FUNCTION SPEED_CONTROL : INT
VAR_INPUT
	ixLevel : INT;
END_VAR

SPEED_CONTROL := (50 - ixLevel) * 10;
IF SPEED_CONTROL < 0 THEN;
	SPEED_CONTROL := 0;
END_IF

END_FUNCTION

(* stored: Version 1.1.0.1
   POU SPEED_CONTROL: Id {2597bb6b-e7d4-4b85-89da-19acc4178c50}, SpecialFunc None *)
